(* IEC 61131-3 sources: tsplc/packages/vscode-extension/tests/fixtures/conveyor/transport/FB_Conveyor/methods/SetMotionSignal, 2 files *)

(* ---- SetMotionSignal.declaration.st ---- *)
METHOD PUBLIC SetMotionSignal
VAR_INPUT
	Asserted : BOOL;
END_VAR
VAR
	ZoneIndex : UINT;
END_VAR

(* ---- SetMotionSignal.implementation.st ---- *)
IF pConveyor = 0 THEN
	RETURN;
END_IF;

IF pConveyor^.ZoneCount > PlantConstants.ZoneCapacity THEN
	RETURN;
END_IF;

FOR ZoneIndex := 1 TO pConveyor^.ZoneCount DO
	pConveyor^.Zones[ZoneIndex].Output.MotionAsserted := Asserted;
END_FOR;
